(* IEC 61131-3 sources: PLC_Gen_Frame/Agents4PLC_release/results/task_1778470003, 1 file *)

(* ---- output.ST ---- *)
FUNCTION_BLOCK in
VAR_INPUT
    ProximitySensor : BOOL;
    ElapsedTime : DINT;
END_VAR
VAR_OUTPUT
    DoorOpen : BOOL;
END_VAR

// Generated by DummyPLCGenerator

END_FUNCTION_BLOCK
